(* IEC 61131-3 sources: plc-st-coding-agent/progress/evidence/full_r8_20261110b/native_evidence/codex_minimax-m27/public-easy-06/0, 1 file *)

(* ---- candidate.st ---- *)
FUNCTION_BLOCK FB
VAR_INPUT
    DO_LOW : BOOL;
    AERATION_E_STOP_NC : BOOL;
END_VAR
VAR_OUTPUT
    BLOWER_RUN : BOOL;
    AERATION_BLOWER_CYCLE_COUNT : UINT;
END_VAR
VAR
    prev_blower_run : BOOL := FALSE;
    delay_counter : UINT := 0;
END_VAR

// Increment cycle count on rising edge of BLOWER_RUN
IF BLOWER_RUN AND NOT prev_blower_run THEN
    AERATION_BLOWER_CYCLE_COUNT := AERATION_BLOWER_CYCLE_COUNT + 1;
END_IF

// Update previous state for next cycle edge detection
prev_blower_run := BLOWER_RUN;

// Check if start conditions are met
IF DO_LOW AND AERATION_E_STOP_NC THEN
    delay_counter := delay_counter + 1;
    IF delay_counter >= 5 THEN
        BLOWER_RUN := TRUE;
    ELSE
        BLOWER_RUN := FALSE;
    END_IF
ELSE
    delay_counter := 0;
    BLOWER_RUN := FALSE;
END_IF
END_FUNCTION_BLOCK
